PROGRAM main
  VAR
    Fill_Btn AT %IX0.0 : BOOL;
    Disch_Btn AT %IX0.1 : BOOL;
    Fill_Valve AT %QX0.0 : BOOL;
    Disch_Valve AT %QX0.1 : BOOL;
    T_Fill : TON;
    T_Disch : TON;
    Fill_Seq : BOOL;
    Disch_Seq : BOOL;
    Fill_Light AT %QX0.2 : BOOL;
    Timer_Disp AT %QW0 : INT;
    Disch_Light AT %QX0.3 : BOOL;
    Fill_sec : LREAL;
    Left_Calc : LREAL;
    Disch_sec : LREAL;
    Fill_Cmd AT %QX0.4 : BOOL;
    Disch_Cmd AT %QX0.5 : BOOL;
    Preset_s AT %MW1 : INT := 10;
    Level AT %MW0 : INT := 0;
    Preset_T : TIME;
    Preset_R : LREAL;
    Preset_R0 : LREAL;
    Step_Lvl : INT;
    Tick : TON;
    Preset_ms : INT;
    Fill_Analog AT %QW1 : INT;
    Disch_Analog AT %QW2 : INT;
    Level_Raw AT %IW0 : INT;
    Tank_Level_Raw AT %MW2 : INT := 0;
  END_VAR
  VAR_EXTERNAL
  END_VAR
  VAR_INPUT
  END_VAR
  VAR  (* added by the conversion: wires and edge detectors of the diagram *)
    _MOVE103_OUT : BOOL;
  END_VAR

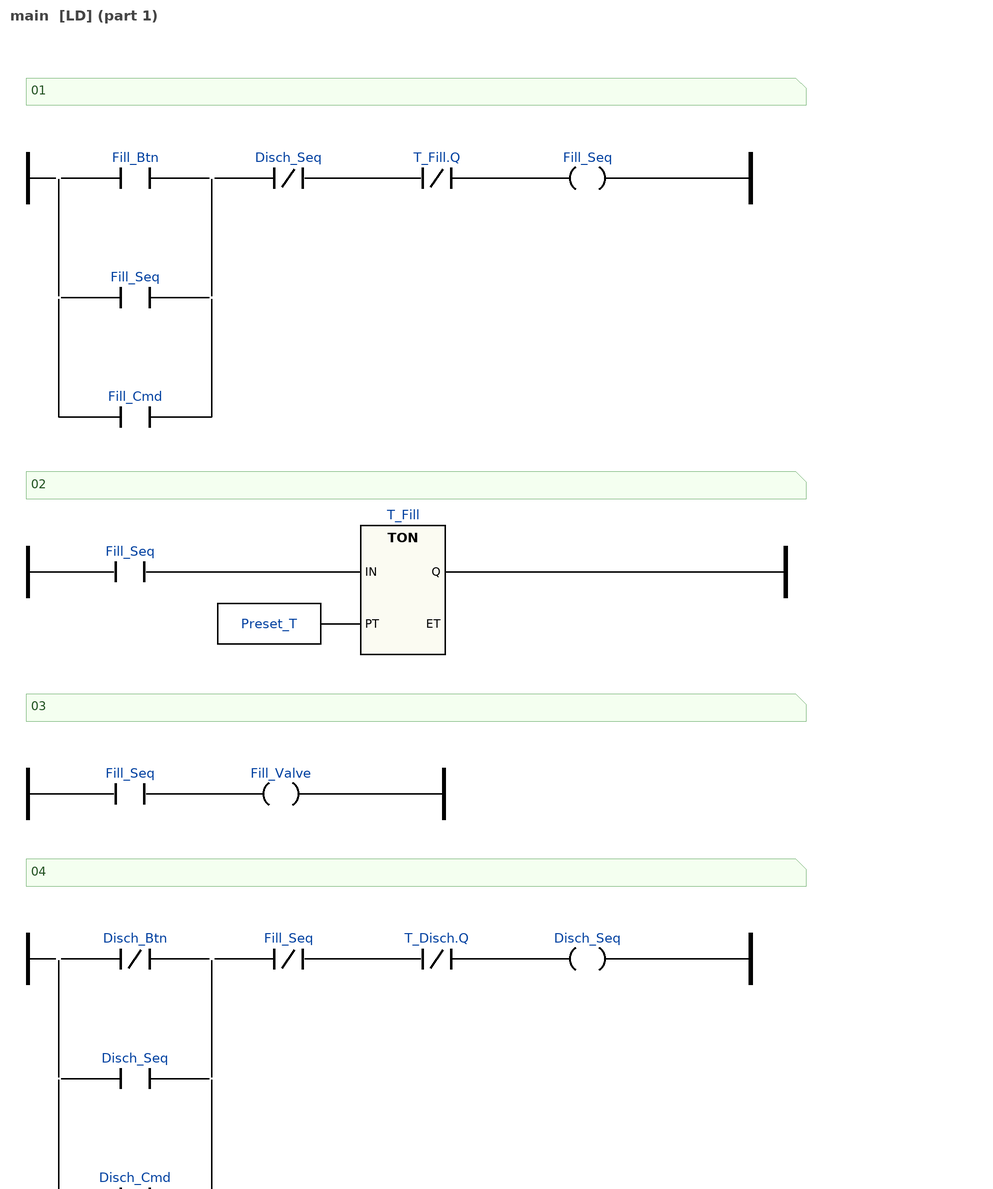
(* LD diagram, written out as Structured Text *)
(* 01 *)
Fill_Seq := (Fill_Btn OR Fill_Seq OR Fill_Cmd) AND NOT Disch_Seq AND NOT T_Fill.Q;
(* 02 *)
(* 03 *)
Fill_Valve := Fill_Seq;
(* 04 *)
Disch_Seq := (NOT Disch_Btn OR Disch_Seq OR Disch_Cmd) AND NOT Fill_Seq AND NOT T_Disch.Q;
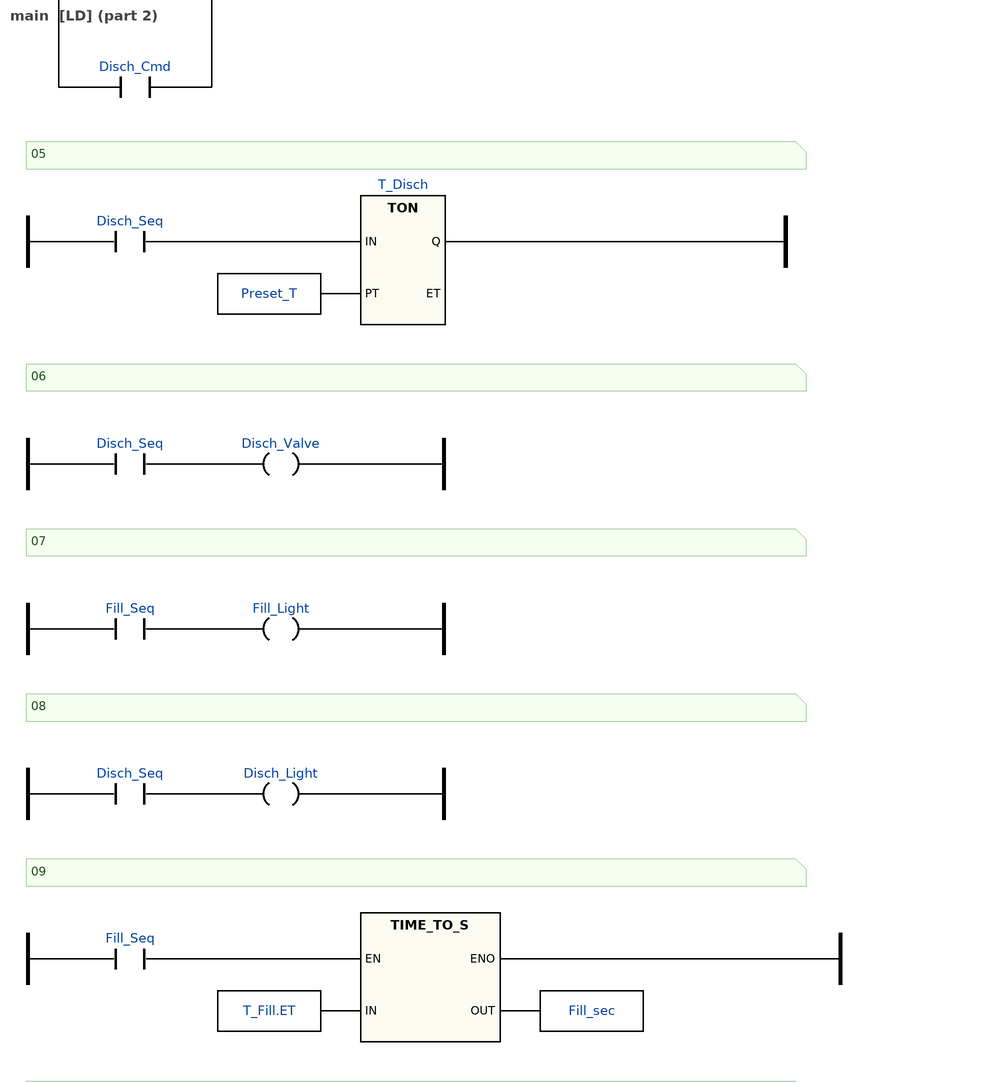
(* 05 *)
(* 06 *)
Disch_Valve := Disch_Seq;
(* 07 *)
Fill_Light := Fill_Seq;
(* 08 *)
Disch_Light := Disch_Seq;
(* 09 *)
IF Fill_Seq THEN Fill_sec := TIME_TO_S(T_Fill.ET); END_IF;
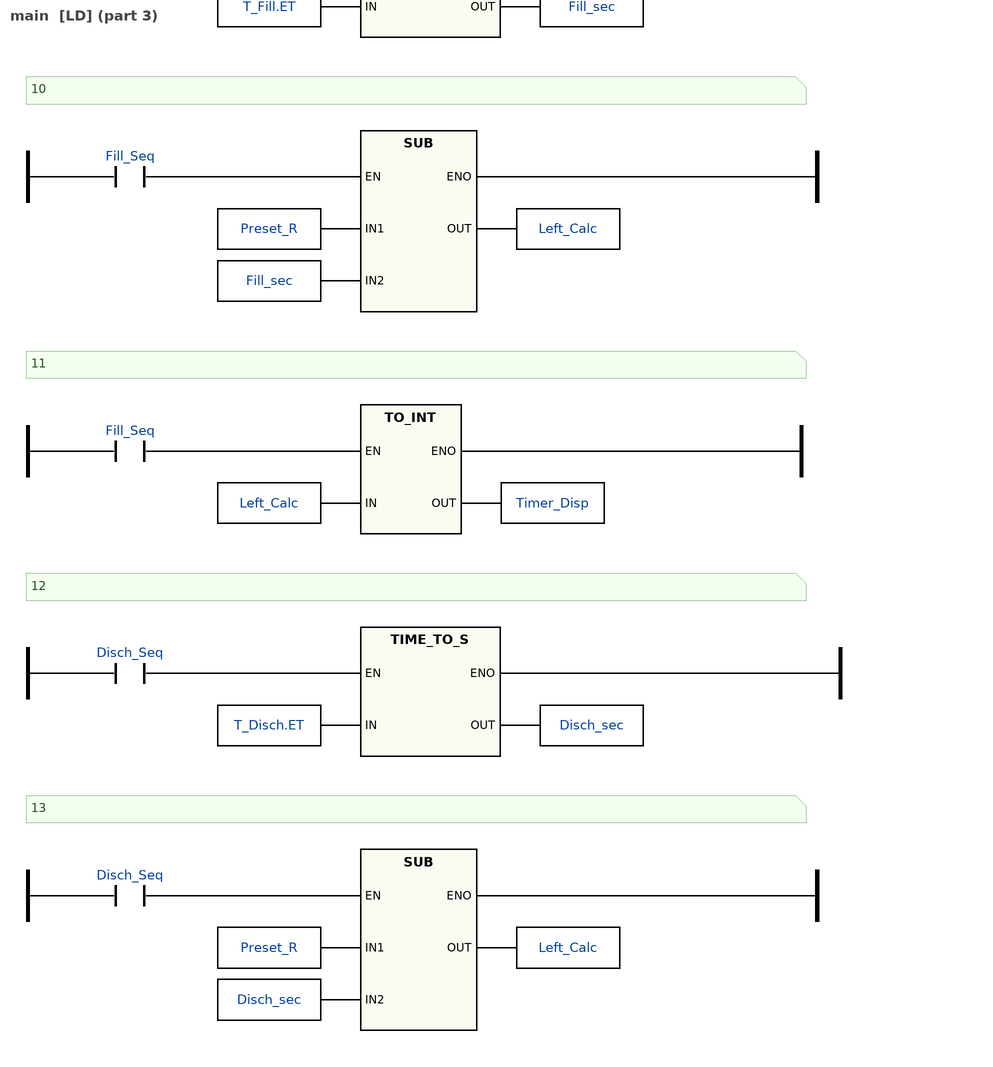
(* 10 *)
IF Fill_Seq THEN Left_Calc := Preset_R - Fill_sec; END_IF;
(* 11 *)
IF Fill_Seq THEN Timer_Disp := TO_INT(Left_Calc); END_IF;
(* 12 *)
IF Disch_Seq THEN Disch_sec := TIME_TO_S(T_Disch.ET); END_IF;
(* 13 *)
IF Disch_Seq THEN Left_Calc := Preset_R - Disch_sec; END_IF;
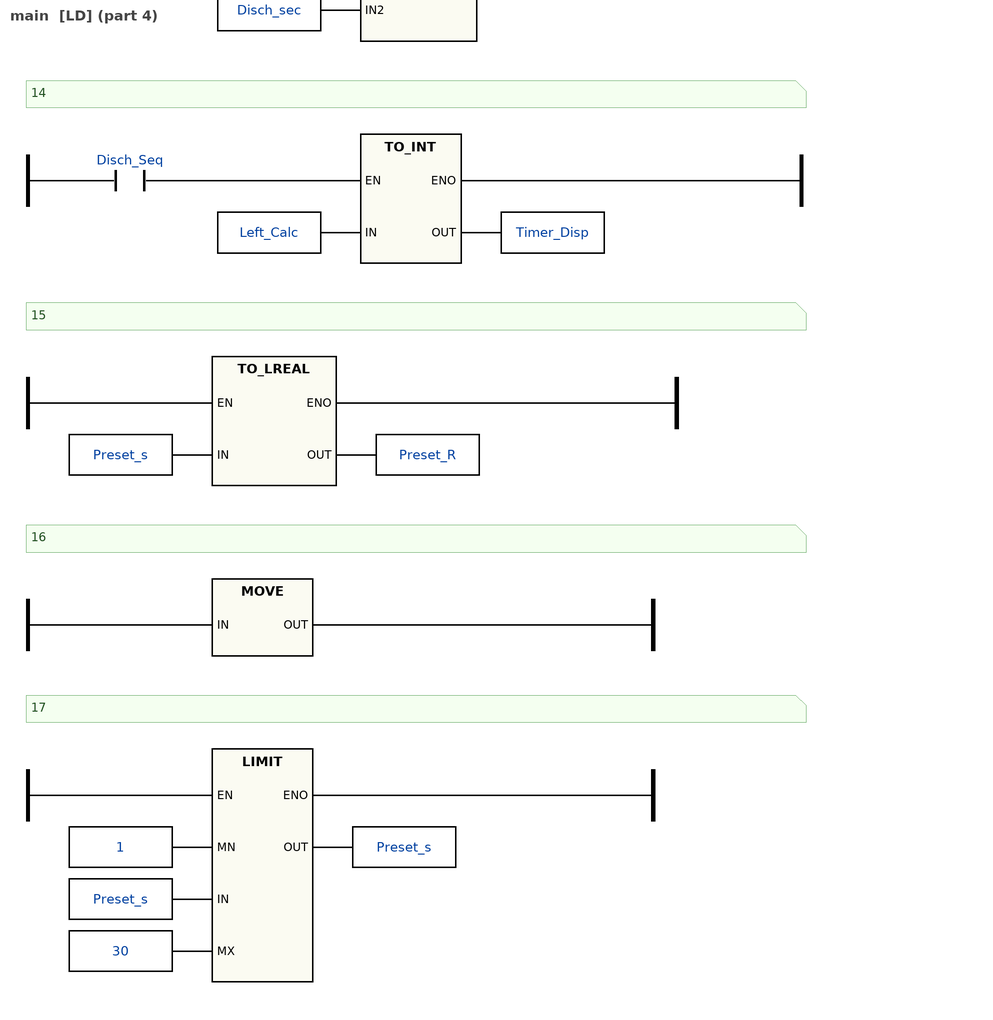
(* 14 *)
IF Disch_Seq THEN Timer_Disp := TO_INT(Left_Calc); END_IF;
(* 15 *)
Preset_R := TO_LREAL(Preset_s);
(* 16 *)
(* 17 *)
Preset_s := LIMIT(1, Preset_s, 30);
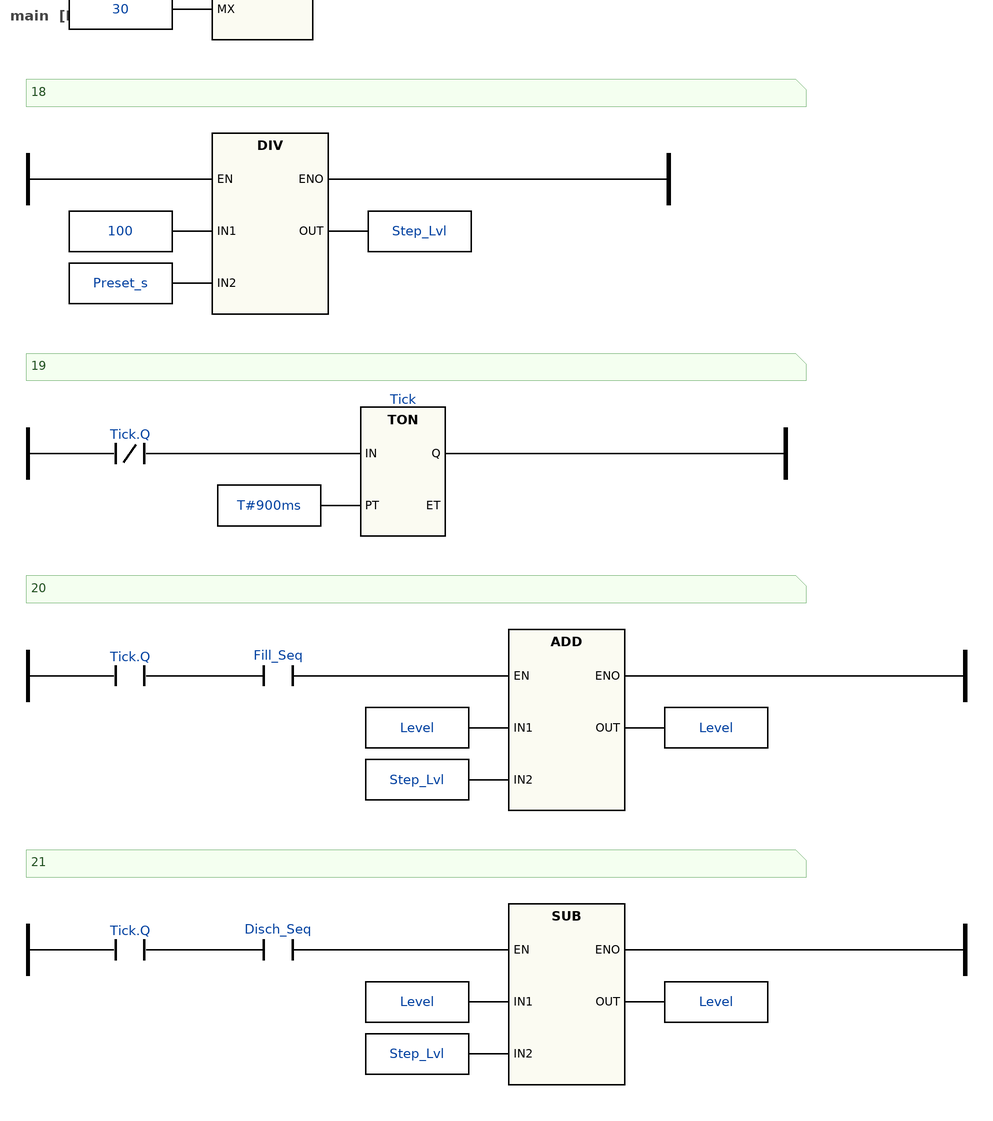
(* 18 *)
Step_Lvl := 100 / Preset_s;
(* 19 *)
(* 20 *)
IF Tick.Q AND Fill_Seq THEN Level := Level + Step_Lvl; END_IF;
(* 21 *)
IF Tick.Q AND Disch_Seq THEN Level := Level - Step_Lvl; END_IF;
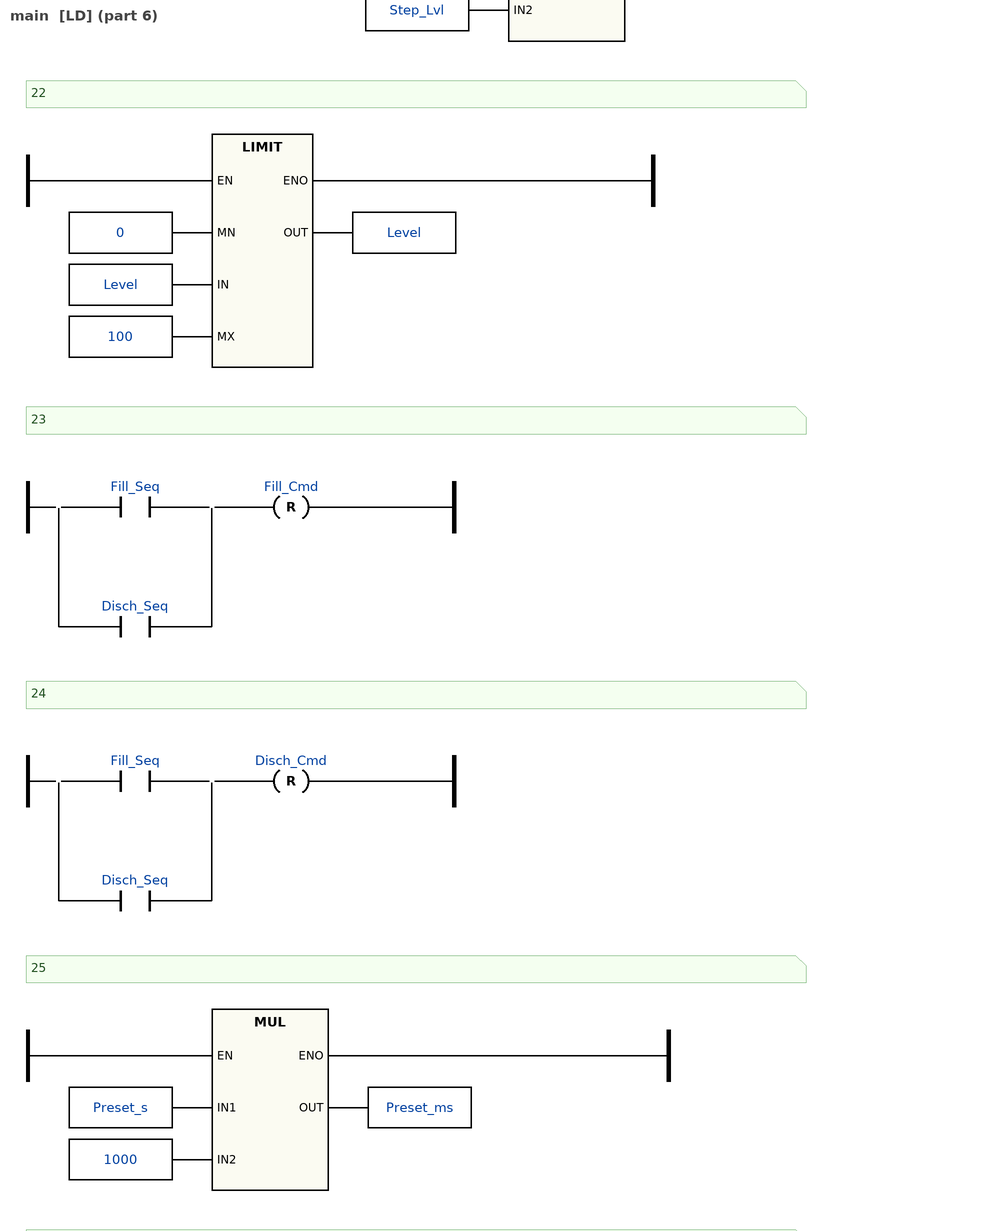
(* 22 *)
Level := LIMIT(0, Level, 100);
(* 23 *)
IF Fill_Seq OR Disch_Seq THEN Fill_Cmd := FALSE; END_IF;
(* 24 *)
IF Fill_Seq OR Disch_Seq THEN Disch_Cmd := FALSE; END_IF;
(* 25 *)
Preset_ms := Preset_s * 1000;
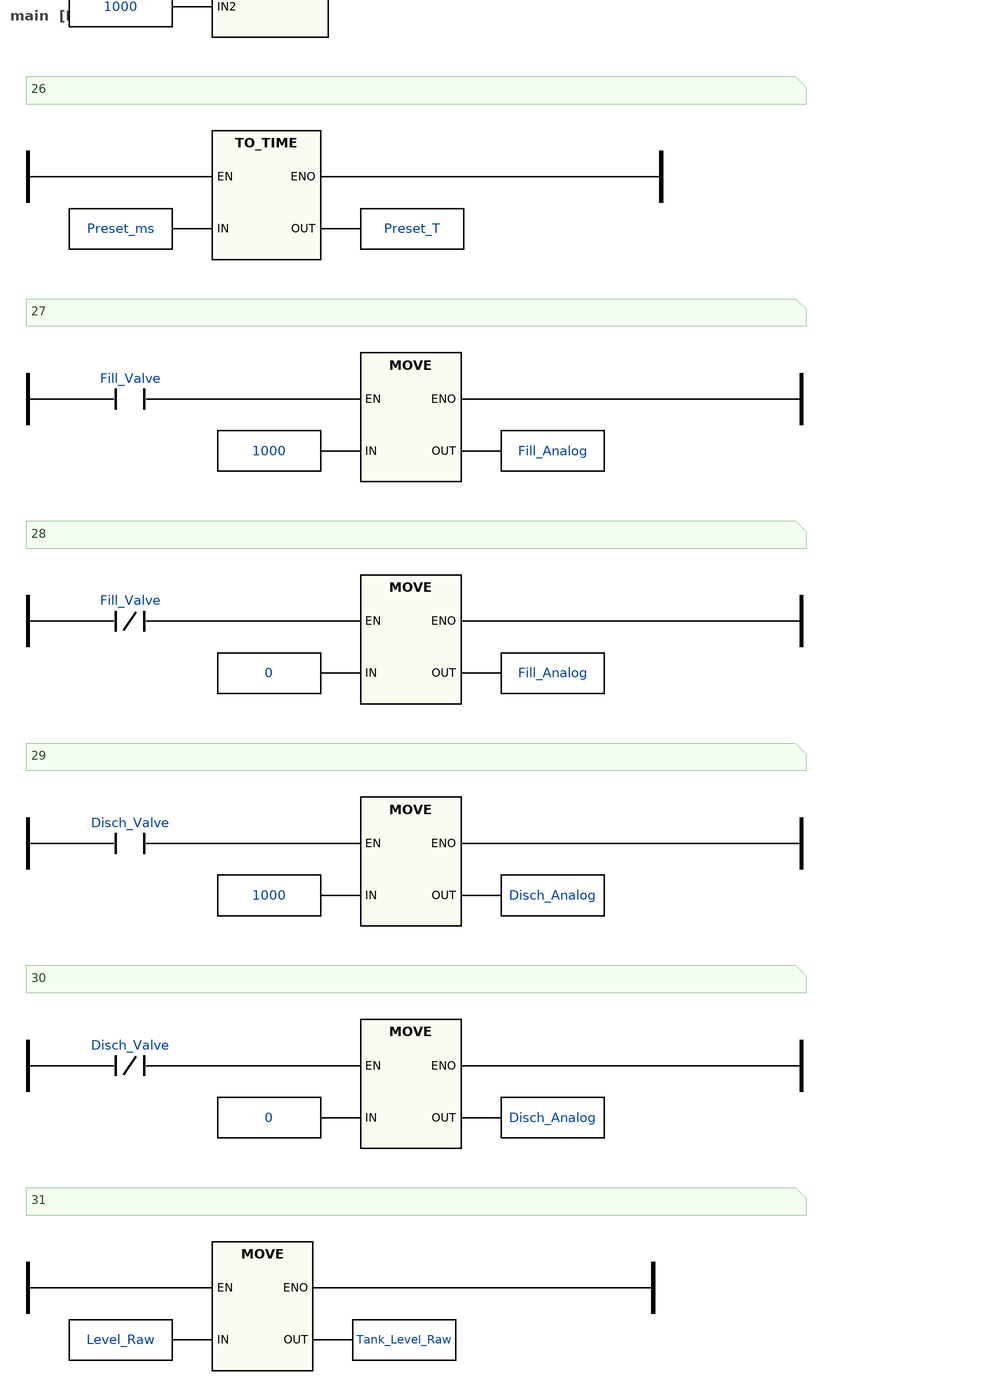
(* 26 *)
Preset_T := TO_TIME(Preset_ms);
(* 27 *)
IF Fill_Valve THEN Fill_Analog := 1000; END_IF;
(* 28 *)
IF NOT Fill_Valve THEN Fill_Analog := 0; END_IF;
(* 29 *)
IF Disch_Valve THEN Disch_Analog := 1000; END_IF;
(* 30 *)
IF NOT Disch_Valve THEN Disch_Analog := 0; END_IF;
(* 31 *)
Tank_Level_Raw := Level_Raw;
T_Fill(IN := Fill_Seq, PT := Preset_T);
T_Disch(IN := Disch_Seq, PT := Preset_T);
_MOVE103_OUT := TRUE;
Tick(IN := NOT Tick.Q, PT := T#900ms);
END_PROGRAM
